(* IEC 61131-3 sources: trust-platform/examples/OSCAT/water_booster_pump_station/non-oop/src, 3 files *)

(* ---- Main.st ---- *)
FUNCTION_BLOCK BoosterStationClassic
VAR
    Pump1Runtime : REAL := REAL#120.0;
    Pump2Runtime : REAL := REAL#20.0;
    Pump3Runtime : REAL := REAL#60.0;
    LeadPumpIdValue : INT;
    RunningPumpCountValue : INT;
    AlarmActiveValue : BOOL;
    AlarmCountValue : INT;
END_VAR

METHOD PUBLIC Update : INT
VAR_INPUT
    StartCommand : BOOL;
    SuctionOk : BOOL;
    Pump1Fault : BOOL;
    Pump2Fault : BOOL;
    Pump3Fault : BOOL;
END_VAR
IF NOT SuctionOk THEN
    AlarmActiveValue := TRUE;
    AlarmCountValue := AlarmCountValue + INT#1;
    LeadPumpIdValue := INT#0;
ELSIF StartCommand THEN
    IF NOT Pump1Fault AND (Pump2Fault OR Pump1Runtime <= Pump2Runtime) AND (Pump3Fault OR Pump1Runtime <= Pump3Runtime) THEN
        LeadPumpIdValue := INT#1;
        RunningPumpCountValue := INT#1;
    ELSIF NOT Pump2Fault AND (Pump3Fault OR Pump2Runtime <= Pump3Runtime) THEN
        LeadPumpIdValue := INT#2;
        RunningPumpCountValue := INT#1;
    ELSIF NOT Pump3Fault THEN
        LeadPumpIdValue := INT#3;
        RunningPumpCountValue := INT#1;
    ELSE
        AlarmActiveValue := TRUE;
        AlarmCountValue := AlarmCountValue + INT#1;
        LeadPumpIdValue := INT#0;
        RunningPumpCountValue := INT#0;
    END_IF;
ELSE
    LeadPumpIdValue := INT#0;
    RunningPumpCountValue := INT#0;
END_IF;
Update := LeadPumpIdValue;
END_METHOD

PUBLIC PROPERTY LeadPumpId : INT
GET
    LeadPumpId := LeadPumpIdValue;
END_GET
END_PROPERTY

PUBLIC PROPERTY RunningPumpCount : INT
GET
    RunningPumpCount := RunningPumpCountValue;
END_GET
END_PROPERTY

PUBLIC PROPERTY AlarmActive : BOOL
GET
    AlarmActive := AlarmActiveValue;
END_GET
END_PROPERTY

PUBLIC PROPERTY AlarmCount : INT
GET
    AlarmCount := AlarmCountValue;
END_GET
END_PROPERTY
END_FUNCTION_BLOCK

PROGRAM Main
VAR
    Station : BoosterStationClassic;
    LeadId : INT;
END_VAR
LeadId := Station.Update(StartCommand := TRUE, SuctionOk := TRUE, Pump1Fault := FALSE, Pump2Fault := FALSE, Pump3Fault := FALSE);
END_PROGRAM

(* ---- Configuration.st ---- *)
CONFIGURATION WaterBoosterClassicConfiguration
RESOURCE WaterBoosterClassic ON PLC
    TASK MainTask (INTERVAL := T#100ms, PRIORITY := 1);
    PROGRAM Station WITH MainTask : Main;
END_RESOURCE
END_CONFIGURATION

(* ---- Tests.st ---- *)
TEST_PROGRAM BoosterClassicSelectsLeadWithDirectBranches
VAR
    Station : BoosterStationClassic;
END_VAR

ASSERT_EQUAL(EXPECTED := INT#2, ACTUAL := Station.Update(StartCommand := TRUE, SuctionOk := TRUE, Pump1Fault := FALSE, Pump2Fault := FALSE, Pump3Fault := FALSE));
ASSERT_EQUAL(EXPECTED := INT#3, ACTUAL := Station.Update(StartCommand := TRUE, SuctionOk := TRUE, Pump1Fault := FALSE, Pump2Fault := TRUE, Pump3Fault := FALSE));
ASSERT_EQUAL(EXPECTED := INT#0, ACTUAL := Station.Update(StartCommand := TRUE, SuctionOk := TRUE, Pump1Fault := TRUE, Pump2Fault := TRUE, Pump3Fault := TRUE));
ASSERT_TRUE(IN := Station.AlarmActive);
ASSERT_EQUAL(EXPECTED := INT#1, ACTUAL := Station.AlarmCount);
END_TEST_PROGRAM
